// TIA Portal V20 export
Screen "USER_OPERATION"  1276x673
  ScreenItem "Move_Legend" at 1184,2 size 90x60  Type=HmiButton
  ScreenItem "Button_Back" at 2,2 size 90x60  Type=HmiButton
  ScreenItem "Fusszeile_Button_ManualOPMode" at 95,2 size 90x60  Type=HmiButton
  ScreenItem "Line_Header_X0_Y64" at 0,64 size 1275x0  Type=HmiLine
  ScreenItem "Line_Header_X0_Y64_1" at 0,64 size 1265x0  Type=HmiLine
  ScreenItem "Title_ScreenOverview_X390_Y2_3" at 384,5 size 510x57  Type=HmiTextBox
  ScreenItem "Move_Legend_1" at 1091,2 size 90x60  Type=HmiButton
  ScreenItem "Line_Header_X0_Y64_2" at 0,64 size 1275x0  Type=HmiLine
  ScreenItem "LSicar_MoveValve_HmiCtrl_1" at 5,64 size 1273x72  Type=HmiFaceplateContainer
  ScreenItem "Line_Header_X0_Y64_3" at 0,64 size 1265x0  Type=HmiLine
  ScreenItem "LSicar_MoveValve_HmiCtrl_6" at 5,446 size 1273x72  Type=HmiFaceplateContainer
  ScreenItem "LSicar_MoveValve_HmiCtrl_7" at 5,523 size 1273x72  Type=HmiFaceplateContainer
  ScreenItem "LSicar_MoveValve_HmiCtrl_8" at 5,601 size 1273x72  Type=HmiFaceplateContainer
  ScreenItem "LSicar_MoveValve_HmiCtrl_2" at 5,138 size 1273x72  Type=HmiFaceplateContainer
  ScreenItem "LSicar_MoveValve_HmiCtrl_3" at 5,215 size 1273x72  Type=HmiFaceplateContainer
  ScreenItem "LSicar_MoveValve_HmiCtrl_4" at 5,292 size 1273x72  Type=HmiFaceplateContainer
  ScreenItem "LSicar_MoveValve_HmiCtrl_5" at 5,369 size 1273x72  Type=HmiFaceplateContainer
  ScreenItem "LSicar_MoveValve_HmiCtrl_9" at 5,64 size 1273x72  Type=HmiFaceplateContainer
  ScreenItem "LSicar_MoveValve_HmiCtrl_14" at 5,446 size 1273x72  Type=HmiFaceplateContainer
  ScreenItem "LSicar_MoveValve_HmiCtrl_15" at 4,522 size 1273x72  Type=HmiFaceplateContainer
  ScreenItem "LSicar_MoveValve_HmiCtrl_16" at 4,599 size 1273x72  Type=HmiFaceplateContainer
  ScreenItem "LSicar_MoveValve_HmiCtrl_10" at 5,136 size 1273x72  Type=HmiFaceplateContainer
  ScreenItem "LSicar_MoveValve_HmiCtrl_11" at 5,214 size 1273x72  Type=HmiFaceplateContainer
  ScreenItem "LSicar_MoveValve_HmiCtrl_12" at 5,292 size 1273x72  Type=HmiFaceplateContainer
  ScreenItem "LSicar_MoveValve_HmiCtrl_13" at 5,370 size 1273x72  Type=HmiFaceplateContainer
